Fanuc KAREL source: NC0072.KL

PROGRAM NC0072
%NOLOCKGROUP
ROUTINE R
VAR
  X : INTEGER
BEGIN
  X = 1
  WHILE X < 2 DO
    X = X + 1
  ENDWHILE
END R
BEGIN
  R
END NC0072
